Fanuc KAREL source: KA00166.KL

PROGRAM KA00166
%NOLOCKGROUP
VAR
  SRC: ARRAY[4] OF BOOLEAN
  DST: ARRAY[4] OF STRING[20]
BEGIN
  DST = SRC
END KA00166
